FUNCTION_BLOCK IOTest16Logic (* Basic Function Block Type *)
  (* Standard: 61499-2 *)
  (* Version 0.0, 11/13/2026, Sandeep Patil, Flexbridge AB, Template *)
  PACKAGE Flexbridge.FestoMPS400;
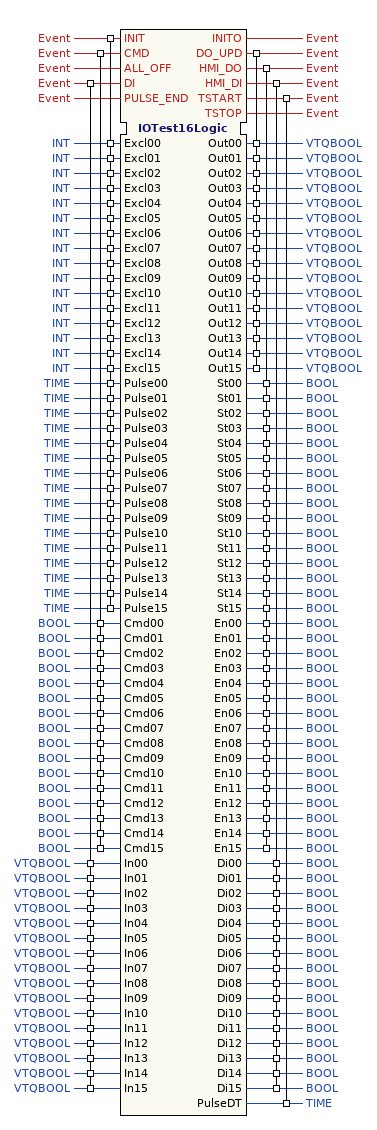
  EVENT_INPUT
    INIT WITH Excl00, Excl01, Excl02, Excl03, Excl04, Excl05, Excl06, Excl07, Excl08, Excl09, Excl10, Excl11, Excl12, Excl13, Excl14, Excl15, Pulse00, Pulse01, Pulse02, Pulse03, Pulse04, Pulse05, Pulse06, Pulse07, Pulse08, Pulse09, Pulse10, Pulse11, Pulse12, Pulse13, Pulse14, Pulse15; (* Initialise; takes over the exclusive pairs and pulse times *)
    CMD WITH Cmd00, Cmd01, Cmd02, Cmd03, Cmd04, Cmd05, Cmd06, Cmd07, Cmd08, Cmd09, Cmd10, Cmd11, Cmd12, Cmd13, Cmd14, Cmd15; (* Button states requested on the HMI *)
    ALL_OFF; (* Switch every output off *)
    DI WITH In00, In01, In02, In03, In04, In05, In06, In07, In08, In09, In10, In11, In12, In13, In14, In15; (* An input channel changed *)
    PULSE_END; (* Pulse timer elapsed *)
  END_EVENT
  EVENT_OUTPUT
    INITO; (* Initialisation done *)
    DO_UPD WITH Out00, Out01, Out02, Out03, Out04, Out05, Out06, Out07, Out08, Out09, Out10, Out11, Out12, Out13, Out14, Out15; (* New output values for the dOSignal blocks *)
    HMI_DO WITH St00, St01, St02, St03, St04, St05, St06, St07, St08, St09, St10, St11, St12, St13, St14, St15, En00, En01, En02, En03, En04, En05, En06, En07, En08, En09, En10, En11, En12, En13, En14, En15; (* Output states and enabled buttons for the HMI *)
    HMI_DI WITH Di00, Di01, Di02, Di03, Di04, Di05, Di06, Di07, Di08, Di09, Di10, Di11, Di12, Di13, Di14, Di15; (* Input values for the HMI *)
    TSTART WITH PulseDT; (* Start the pulse timer *)
    TSTOP; (* Cancel the pulse timer *)
  END_EVENT
  VAR_INPUT
    Excl00 : INT := -1; (* Output that must never be on together with output 00; -1 = none *)
    Excl01 : INT := -1; (* Output that must never be on together with output 01; -1 = none *)
    Excl02 : INT := -1; (* Output that must never be on together with output 02; -1 = none *)
    Excl03 : INT := -1; (* Output that must never be on together with output 03; -1 = none *)
    Excl04 : INT := -1; (* Output that must never be on together with output 04; -1 = none *)
    Excl05 : INT := -1; (* Output that must never be on together with output 05; -1 = none *)
    Excl06 : INT := -1; (* Output that must never be on together with output 06; -1 = none *)
    Excl07 : INT := -1; (* Output that must never be on together with output 07; -1 = none *)
    Excl08 : INT := -1; (* Output that must never be on together with output 08; -1 = none *)
    Excl09 : INT := -1; (* Output that must never be on together with output 09; -1 = none *)
    Excl10 : INT := -1; (* Output that must never be on together with output 10; -1 = none *)
    Excl11 : INT := -1; (* Output that must never be on together with output 11; -1 = none *)
    Excl12 : INT := -1; (* Output that must never be on together with output 12; -1 = none *)
    Excl13 : INT := -1; (* Output that must never be on together with output 13; -1 = none *)
    Excl14 : INT := -1; (* Output that must never be on together with output 14; -1 = none *)
    Excl15 : INT := -1; (* Output that must never be on together with output 15; -1 = none *)
    Pulse00 : TIME := T#0s; (* Pulse time of output 00; T#0s = toggle *)
    Pulse01 : TIME := T#0s; (* Pulse time of output 01; T#0s = toggle *)
    Pulse02 : TIME := T#0s; (* Pulse time of output 02; T#0s = toggle *)
    Pulse03 : TIME := T#0s; (* Pulse time of output 03; T#0s = toggle *)
    Pulse04 : TIME := T#0s; (* Pulse time of output 04; T#0s = toggle *)
    Pulse05 : TIME := T#0s; (* Pulse time of output 05; T#0s = toggle *)
    Pulse06 : TIME := T#0s; (* Pulse time of output 06; T#0s = toggle *)
    Pulse07 : TIME := T#0s; (* Pulse time of output 07; T#0s = toggle *)
    Pulse08 : TIME := T#0s; (* Pulse time of output 08; T#0s = toggle *)
    Pulse09 : TIME := T#0s; (* Pulse time of output 09; T#0s = toggle *)
    Pulse10 : TIME := T#0s; (* Pulse time of output 10; T#0s = toggle *)
    Pulse11 : TIME := T#0s; (* Pulse time of output 11; T#0s = toggle *)
    Pulse12 : TIME := T#0s; (* Pulse time of output 12; T#0s = toggle *)
    Pulse13 : TIME := T#0s; (* Pulse time of output 13; T#0s = toggle *)
    Pulse14 : TIME := T#0s; (* Pulse time of output 14; T#0s = toggle *)
    Pulse15 : TIME := T#0s; (* Pulse time of output 15; T#0s = toggle *)
    Cmd00 : BOOL; (* Requested state of output 00 *)
    Cmd01 : BOOL; (* Requested state of output 01 *)
    Cmd02 : BOOL; (* Requested state of output 02 *)
    Cmd03 : BOOL; (* Requested state of output 03 *)
    Cmd04 : BOOL; (* Requested state of output 04 *)
    Cmd05 : BOOL; (* Requested state of output 05 *)
    Cmd06 : BOOL; (* Requested state of output 06 *)
    Cmd07 : BOOL; (* Requested state of output 07 *)
    Cmd08 : BOOL; (* Requested state of output 08 *)
    Cmd09 : BOOL; (* Requested state of output 09 *)
    Cmd10 : BOOL; (* Requested state of output 10 *)
    Cmd11 : BOOL; (* Requested state of output 11 *)
    Cmd12 : BOOL; (* Requested state of output 12 *)
    Cmd13 : BOOL; (* Requested state of output 13 *)
    Cmd14 : BOOL; (* Requested state of output 14 *)
    Cmd15 : BOOL; (* Requested state of output 15 *)
    In00 : VTQBOOL; (* Input channel 00 *)
    In01 : VTQBOOL; (* Input channel 01 *)
    In02 : VTQBOOL; (* Input channel 02 *)
    In03 : VTQBOOL; (* Input channel 03 *)
    In04 : VTQBOOL; (* Input channel 04 *)
    In05 : VTQBOOL; (* Input channel 05 *)
    In06 : VTQBOOL; (* Input channel 06 *)
    In07 : VTQBOOL; (* Input channel 07 *)
    In08 : VTQBOOL; (* Input channel 08 *)
    In09 : VTQBOOL; (* Input channel 09 *)
    In10 : VTQBOOL; (* Input channel 10 *)
    In11 : VTQBOOL; (* Input channel 11 *)
    In12 : VTQBOOL; (* Input channel 12 *)
    In13 : VTQBOOL; (* Input channel 13 *)
    In14 : VTQBOOL; (* Input channel 14 *)
    In15 : VTQBOOL; (* Input channel 15 *)
  END_VAR
  VAR_OUTPUT
    Out00 : VTQBOOL; (* Output channel 00 *)
    Out01 : VTQBOOL; (* Output channel 01 *)
    Out02 : VTQBOOL; (* Output channel 02 *)
    Out03 : VTQBOOL; (* Output channel 03 *)
    Out04 : VTQBOOL; (* Output channel 04 *)
    Out05 : VTQBOOL; (* Output channel 05 *)
    Out06 : VTQBOOL; (* Output channel 06 *)
    Out07 : VTQBOOL; (* Output channel 07 *)
    Out08 : VTQBOOL; (* Output channel 08 *)
    Out09 : VTQBOOL; (* Output channel 09 *)
    Out10 : VTQBOOL; (* Output channel 10 *)
    Out11 : VTQBOOL; (* Output channel 11 *)
    Out12 : VTQBOOL; (* Output channel 12 *)
    Out13 : VTQBOOL; (* Output channel 13 *)
    Out14 : VTQBOOL; (* Output channel 14 *)
    Out15 : VTQBOOL; (* Output channel 15 *)
    St00 : BOOL; (* Current state of output 00 *)
    St01 : BOOL; (* Current state of output 01 *)
    St02 : BOOL; (* Current state of output 02 *)
    St03 : BOOL; (* Current state of output 03 *)
    St04 : BOOL; (* Current state of output 04 *)
    St05 : BOOL; (* Current state of output 05 *)
    St06 : BOOL; (* Current state of output 06 *)
    St07 : BOOL; (* Current state of output 07 *)
    St08 : BOOL; (* Current state of output 08 *)
    St09 : BOOL; (* Current state of output 09 *)
    St10 : BOOL; (* Current state of output 10 *)
    St11 : BOOL; (* Current state of output 11 *)
    St12 : BOOL; (* Current state of output 12 *)
    St13 : BOOL; (* Current state of output 13 *)
    St14 : BOOL; (* Current state of output 14 *)
    St15 : BOOL; (* Current state of output 15 *)
    En00 : BOOL; (* Button of output 00 may be pressed *)
    En01 : BOOL; (* Button of output 01 may be pressed *)
    En02 : BOOL; (* Button of output 02 may be pressed *)
    En03 : BOOL; (* Button of output 03 may be pressed *)
    En04 : BOOL; (* Button of output 04 may be pressed *)
    En05 : BOOL; (* Button of output 05 may be pressed *)
    En06 : BOOL; (* Button of output 06 may be pressed *)
    En07 : BOOL; (* Button of output 07 may be pressed *)
    En08 : BOOL; (* Button of output 08 may be pressed *)
    En09 : BOOL; (* Button of output 09 may be pressed *)
    En10 : BOOL; (* Button of output 10 may be pressed *)
    En11 : BOOL; (* Button of output 11 may be pressed *)
    En12 : BOOL; (* Button of output 12 may be pressed *)
    En13 : BOOL; (* Button of output 13 may be pressed *)
    En14 : BOOL; (* Button of output 14 may be pressed *)
    En15 : BOOL; (* Button of output 15 may be pressed *)
    Di00 : BOOL; (* Value of input 00 *)
    Di01 : BOOL; (* Value of input 01 *)
    Di02 : BOOL; (* Value of input 02 *)
    Di03 : BOOL; (* Value of input 03 *)
    Di04 : BOOL; (* Value of input 04 *)
    Di05 : BOOL; (* Value of input 05 *)
    Di06 : BOOL; (* Value of input 06 *)
    Di07 : BOOL; (* Value of input 07 *)
    Di08 : BOOL; (* Value of input 08 *)
    Di09 : BOOL; (* Value of input 09 *)
    Di10 : BOOL; (* Value of input 10 *)
    Di11 : BOOL; (* Value of input 11 *)
    Di12 : BOOL; (* Value of input 12 *)
    Di13 : BOOL; (* Value of input 13 *)
    Di14 : BOOL; (* Value of input 14 *)
    Di15 : BOOL; (* Value of input 15 *)
    PulseDT : TIME; (* Duration of the pulse being started *)
  END_VAR
  VAR
    Changed : BOOL; (* An output state changed *)
    StartPulse : BOOL; (* A pulse timer must be started *)
    StopPulse : BOOL; (* The pulse timer must be cancelled *)
    PulseCh : INT := -1; (* Output whose pulse is running; -1 = none *)
    PrevRq00 : BOOL; (* Last requested state of output 00 *)
    PrevRq01 : BOOL; (* Last requested state of output 01 *)
    PrevRq02 : BOOL; (* Last requested state of output 02 *)
    PrevRq03 : BOOL; (* Last requested state of output 03 *)
    PrevRq04 : BOOL; (* Last requested state of output 04 *)
    PrevRq05 : BOOL; (* Last requested state of output 05 *)
    PrevRq06 : BOOL; (* Last requested state of output 06 *)
    PrevRq07 : BOOL; (* Last requested state of output 07 *)
    PrevRq08 : BOOL; (* Last requested state of output 08 *)
    PrevRq09 : BOOL; (* Last requested state of output 09 *)
    PrevRq10 : BOOL; (* Last requested state of output 10 *)
    PrevRq11 : BOOL; (* Last requested state of output 11 *)
    PrevRq12 : BOOL; (* Last requested state of output 12 *)
    PrevRq13 : BOOL; (* Last requested state of output 13 *)
    PrevRq14 : BOOL; (* Last requested state of output 14 *)
    PrevRq15 : BOOL; (* Last requested state of output 15 *)
  END_VAR
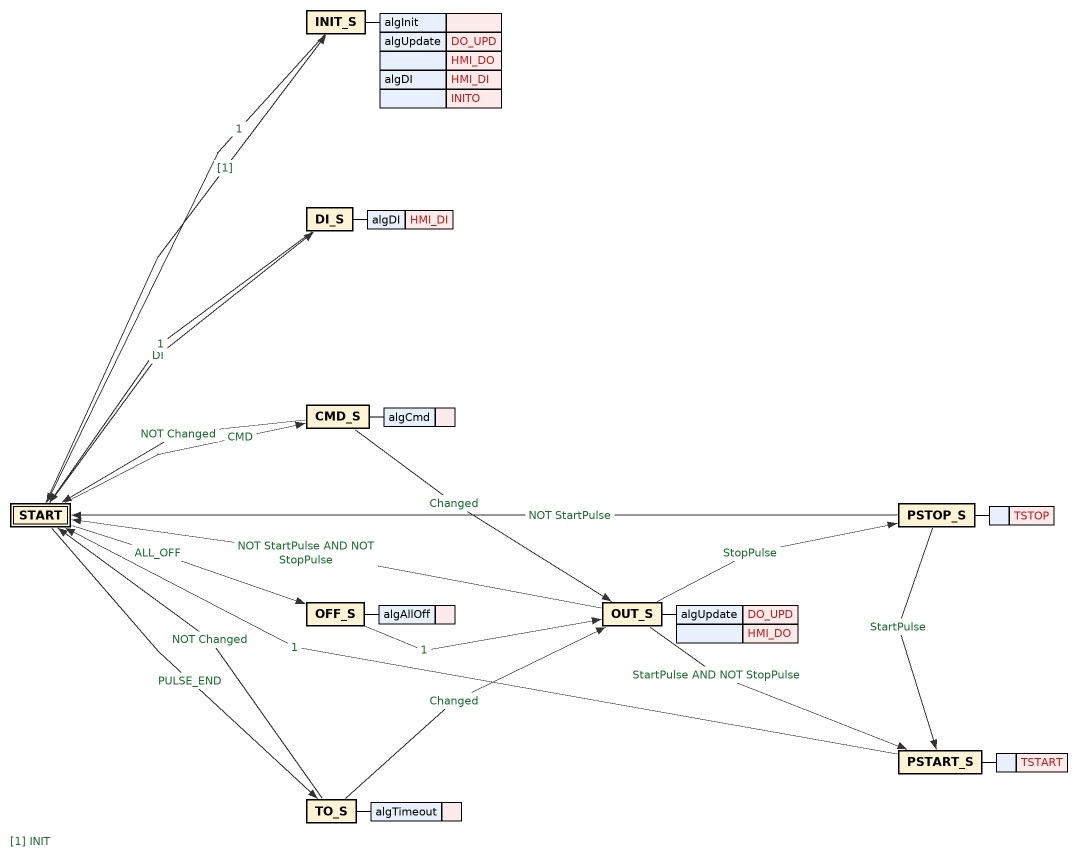
  EC_STATES
    START; (* Initial State *)
    INIT_S : algInit, algUpdate -> DO_UPD, -> HMI_DO, algDI -> HMI_DI, -> INITO;
    DI_S : algDI -> HMI_DI;
    CMD_S : algCmd;
    OFF_S : algAllOff;
    TO_S : algTimeout;
    OUT_S : algUpdate -> DO_UPD, -> HMI_DO;
    PSTOP_S : -> TSTOP;
    PSTART_S : -> TSTART;
  END_STATES
  EC_TRANSITIONS
    START TO INIT_S := INIT;
    INIT_S TO START := 1;
    START TO DI_S := DI;
    DI_S TO START := 1;
    START TO CMD_S := CMD;
    CMD_S TO OUT_S := Changed;
    CMD_S TO START := NOT Changed;
    START TO OFF_S := ALL_OFF;
    OFF_S TO OUT_S := 1;
    START TO TO_S := PULSE_END;
    TO_S TO OUT_S := Changed;
    TO_S TO START := NOT Changed;
    OUT_S TO PSTOP_S := StopPulse;
    OUT_S TO PSTART_S := StartPulse AND NOT StopPulse;
    OUT_S TO START := NOT StartPulse AND NOT StopPulse;
    PSTOP_S TO PSTART_S := StartPulse;
    PSTOP_S TO START := NOT StartPulse;
    PSTART_S TO START := 1;
  END_TRANSITIONS
  ALGORITHM algInit IN ST:
(* All outputs off, no pulse running *)
St00 := FALSE;
PrevRq00 := FALSE;
St01 := FALSE;
PrevRq01 := FALSE;
St02 := FALSE;
PrevRq02 := FALSE;
St03 := FALSE;
PrevRq03 := FALSE;
St04 := FALSE;
PrevRq04 := FALSE;
St05 := FALSE;
PrevRq05 := FALSE;
St06 := FALSE;
PrevRq06 := FALSE;
St07 := FALSE;
PrevRq07 := FALSE;
St08 := FALSE;
PrevRq08 := FALSE;
St09 := FALSE;
PrevRq09 := FALSE;
St10 := FALSE;
PrevRq10 := FALSE;
St11 := FALSE;
PrevRq11 := FALSE;
St12 := FALSE;
PrevRq12 := FALSE;
St13 := FALSE;
PrevRq13 := FALSE;
St14 := FALSE;
PrevRq14 := FALSE;
St15 := FALSE;
PrevRq15 := FALSE;
PulseCh := -1;
Changed := FALSE;
StartPulse := FALSE;
StopPulse := FALSE;
  END_ALGORITHM
  ALGORITHM algDI IN ST:
(* Copy the input values for the HMI *)
Di00 := In00.value;
Di01 := In01.value;
Di02 := In02.value;
Di03 := In03.value;
Di04 := In04.value;
Di05 := In05.value;
Di06 := In06.value;
Di07 := In07.value;
Di08 := In08.value;
Di09 := In09.value;
Di10 := In10.value;
Di11 := In11.value;
Di12 := In12.value;
Di13 := In13.value;
Di14 := In14.value;
Di15 := In15.value;
  END_ALGORITHM
  ALGORITHM algCmd IN ST:
VAR
  aSt : ARRAY[0..15] OF BOOL;
  aRq : ARRAY[0..15] OF BOOL;
  aPr : ARRAY[0..15] OF BOOL;
  aEx : ARRAY[0..15] OF INT;
  aPu : ARRAY[0..15] OF TIME;
  i : INT;
  p : INT;
  allowed : BOOL;
END_VAR
aSt[0] := St00;
aSt[1] := St01;
aSt[2] := St02;
aSt[3] := St03;
aSt[4] := St04;
aSt[5] := St05;
aSt[6] := St06;
aSt[7] := St07;
aSt[8] := St08;
aSt[9] := St09;
aSt[10] := St10;
aSt[11] := St11;
aSt[12] := St12;
aSt[13] := St13;
aSt[14] := St14;
aSt[15] := St15;
aRq[0] := Cmd00;
aRq[1] := Cmd01;
aRq[2] := Cmd02;
aRq[3] := Cmd03;
aRq[4] := Cmd04;
aRq[5] := Cmd05;
aRq[6] := Cmd06;
aRq[7] := Cmd07;
aRq[8] := Cmd08;
aRq[9] := Cmd09;
aRq[10] := Cmd10;
aRq[11] := Cmd11;
aRq[12] := Cmd12;
aRq[13] := Cmd13;
aRq[14] := Cmd14;
aRq[15] := Cmd15;
aPr[0] := PrevRq00;
aPr[1] := PrevRq01;
aPr[2] := PrevRq02;
aPr[3] := PrevRq03;
aPr[4] := PrevRq04;
aPr[5] := PrevRq05;
aPr[6] := PrevRq06;
aPr[7] := PrevRq07;
aPr[8] := PrevRq08;
aPr[9] := PrevRq09;
aPr[10] := PrevRq10;
aPr[11] := PrevRq11;
aPr[12] := PrevRq12;
aPr[13] := PrevRq13;
aPr[14] := PrevRq14;
aPr[15] := PrevRq15;
aEx[0] := Excl00;
aEx[1] := Excl01;
aEx[2] := Excl02;
aEx[3] := Excl03;
aEx[4] := Excl04;
aEx[5] := Excl05;
aEx[6] := Excl06;
aEx[7] := Excl07;
aEx[8] := Excl08;
aEx[9] := Excl09;
aEx[10] := Excl10;
aEx[11] := Excl11;
aEx[12] := Excl12;
aEx[13] := Excl13;
aEx[14] := Excl14;
aEx[15] := Excl15;
aPu[0] := Pulse00;
aPu[1] := Pulse01;
aPu[2] := Pulse02;
aPu[3] := Pulse03;
aPu[4] := Pulse04;
aPu[5] := Pulse05;
aPu[6] := Pulse06;
aPu[7] := Pulse07;
aPu[8] := Pulse08;
aPu[9] := Pulse09;
aPu[10] := Pulse10;
aPu[11] := Pulse11;
aPu[12] := Pulse12;
aPu[13] := Pulse13;
aPu[14] := Pulse14;
aPu[15] := Pulse15;
Changed := FALSE;
StartPulse := FALSE;
StopPulse := FALSE;
(* Only buttons whose request changed since the last CMD are handled, so a request that was
   refused earlier never switches an output on later by surprise. *)
FOR i := 0 TO 15 DO
  IF aRq[i] <> aPr[i] THEN
    aPr[i] := aRq[i];
    IF aRq[i] <> aSt[i] THEN
      IF NOT aRq[i] THEN
        (* Switching off is always allowed *)
        aSt[i] := FALSE;
        Changed := TRUE;
        IF PulseCh = i THEN
          PulseCh := -1;
          StopPulse := TRUE;
        END_IF;
      ELSE
        (* Switching on: refused while the partner output is on, or while another pulse runs *)
        allowed := TRUE;
        p := aEx[i];
        IF (p >= 0) AND (p <= 15) THEN
          IF aSt[p] THEN
            allowed := FALSE;
          END_IF;
        END_IF;
        IF (aPu[i] > T#0s) AND (PulseCh >= 0) THEN
          allowed := FALSE;
        END_IF;
        IF allowed THEN
          aSt[i] := TRUE;
          Changed := TRUE;
          IF aPu[i] > T#0s THEN
            PulseCh := i;
            PulseDT := aPu[i];
            StartPulse := TRUE;
          END_IF;
        END_IF;
      END_IF;
    END_IF;
  END_IF;
END_FOR;
St00 := aSt[0];
St01 := aSt[1];
St02 := aSt[2];
St03 := aSt[3];
St04 := aSt[4];
St05 := aSt[5];
St06 := aSt[6];
St07 := aSt[7];
St08 := aSt[8];
St09 := aSt[9];
St10 := aSt[10];
St11 := aSt[11];
St12 := aSt[12];
St13 := aSt[13];
St14 := aSt[14];
St15 := aSt[15];
PrevRq00 := aPr[0];
PrevRq01 := aPr[1];
PrevRq02 := aPr[2];
PrevRq03 := aPr[3];
PrevRq04 := aPr[4];
PrevRq05 := aPr[5];
PrevRq06 := aPr[6];
PrevRq07 := aPr[7];
PrevRq08 := aPr[8];
PrevRq09 := aPr[9];
PrevRq10 := aPr[10];
PrevRq11 := aPr[11];
PrevRq12 := aPr[12];
PrevRq13 := aPr[13];
PrevRq14 := aPr[14];
PrevRq15 := aPr[15];
  END_ALGORITHM
  ALGORITHM algAllOff IN ST:
(* Switch everything off and cancel a running pulse *)
St00 := FALSE;
St01 := FALSE;
St02 := FALSE;
St03 := FALSE;
St04 := FALSE;
St05 := FALSE;
St06 := FALSE;
St07 := FALSE;
St08 := FALSE;
St09 := FALSE;
St10 := FALSE;
St11 := FALSE;
St12 := FALSE;
St13 := FALSE;
St14 := FALSE;
St15 := FALSE;
StopPulse := (PulseCh >= 0);
PulseCh := -1;
StartPulse := FALSE;
Changed := TRUE;
  END_ALGORITHM
  ALGORITHM algTimeout IN ST:
VAR
  aSt : ARRAY[0..15] OF BOOL;
END_VAR
aSt[0] := St00;
aSt[1] := St01;
aSt[2] := St02;
aSt[3] := St03;
aSt[4] := St04;
aSt[5] := St05;
aSt[6] := St06;
aSt[7] := St07;
aSt[8] := St08;
aSt[9] := St09;
aSt[10] := St10;
aSt[11] := St11;
aSt[12] := St12;
aSt[13] := St13;
aSt[14] := St14;
aSt[15] := St15;
Changed := FALSE;
StartPulse := FALSE;
StopPulse := FALSE;
IF (PulseCh >= 0) AND (PulseCh <= 15) THEN
  aSt[PulseCh] := FALSE;
  PulseCh := -1;
  Changed := TRUE;
END_IF;
St00 := aSt[0];
St01 := aSt[1];
St02 := aSt[2];
St03 := aSt[3];
St04 := aSt[4];
St05 := aSt[5];
St06 := aSt[6];
St07 := aSt[7];
St08 := aSt[8];
St09 := aSt[9];
St10 := aSt[10];
St11 := aSt[11];
St12 := aSt[12];
St13 := aSt[13];
St14 := aSt[14];
St15 := aSt[15];
  END_ALGORITHM
  ALGORITHM algUpdate IN ST:
VAR
  aSt : ARRAY[0..15] OF BOOL;
  aEx : ARRAY[0..15] OF INT;
  aPu : ARRAY[0..15] OF TIME;
  aEn : ARRAY[0..15] OF BOOL;
  i : INT;
  p : INT;
END_VAR
aSt[0] := St00;
aSt[1] := St01;
aSt[2] := St02;
aSt[3] := St03;
aSt[4] := St04;
aSt[5] := St05;
aSt[6] := St06;
aSt[7] := St07;
aSt[8] := St08;
aSt[9] := St09;
aSt[10] := St10;
aSt[11] := St11;
aSt[12] := St12;
aSt[13] := St13;
aSt[14] := St14;
aSt[15] := St15;
aEx[0] := Excl00;
aEx[1] := Excl01;
aEx[2] := Excl02;
aEx[3] := Excl03;
aEx[4] := Excl04;
aEx[5] := Excl05;
aEx[6] := Excl06;
aEx[7] := Excl07;
aEx[8] := Excl08;
aEx[9] := Excl09;
aEx[10] := Excl10;
aEx[11] := Excl11;
aEx[12] := Excl12;
aEx[13] := Excl13;
aEx[14] := Excl14;
aEx[15] := Excl15;
aPu[0] := Pulse00;
aPu[1] := Pulse01;
aPu[2] := Pulse02;
aPu[3] := Pulse03;
aPu[4] := Pulse04;
aPu[5] := Pulse05;
aPu[6] := Pulse06;
aPu[7] := Pulse07;
aPu[8] := Pulse08;
aPu[9] := Pulse09;
aPu[10] := Pulse10;
aPu[11] := Pulse11;
aPu[12] := Pulse12;
aPu[13] := Pulse13;
aPu[14] := Pulse14;
aPu[15] := Pulse15;
(* A button is enabled unless its partner output is on, or it is a pulse output while another pulse runs *)
FOR i := 0 TO 15 DO
  aEn[i] := TRUE;
  p := aEx[i];
  IF (p >= 0) AND (p <= 15) THEN
    IF aSt[p] THEN
      aEn[i] := FALSE;
    END_IF;
  END_IF;
  IF (aPu[i] > T#0s) AND (PulseCh >= 0) AND (PulseCh <> i) THEN
    aEn[i] := FALSE;
  END_IF;
END_FOR;
En00 := aEn[0];
En01 := aEn[1];
En02 := aEn[2];
En03 := aEn[3];
En04 := aEn[4];
En05 := aEn[5];
En06 := aEn[6];
En07 := aEn[7];
En08 := aEn[8];
En09 := aEn[9];
En10 := aEn[10];
En11 := aEn[11];
En12 := aEn[12];
En13 := aEn[13];
En14 := aEn[14];
En15 := aEn[15];
Out00.value := St00;
Out01.value := St01;
Out02.value := St02;
Out03.value := St03;
Out04.value := St04;
Out05.value := St05;
Out06.value := St06;
Out07.value := St07;
Out08.value := St08;
Out09.value := St09;
Out10.value := St10;
Out11.value := St11;
Out12.value := St12;
Out13.value := St13;
Out14.value := St14;
Out15.value := St15;
  END_ALGORITHM
END_FUNCTION_BLOCK
